(* IEC 61131-3 sources: kns-port-domestic/upstream/plc-process-lib/src/POUs/Control/FB_PID, 12 files *)

(* ---- FB_PID.decl.st ---- *)
// Назначение: ПИД-регулятор в идеальной форме (Kp, Ti, Td): D по измерению с фильтром первого
//             порядка, anti-windup обратным расчётом с постоянной слежения Tt (по своему выходу
//             или по фактическому выходу механизма rOutAct_pct), пределы и ограничение скорости
//             выхода, Manual и слежение (xTrack) с безударным переходом, внешнее или операторское
//             задание с рампой, прямое и обратное действие, зона нечувствительности, расчёт по
//             реальному dt источника времени и период расчёта tSample, реакция на недостоверную PV.
//             Внутреннее состояние (I, D, PV прошлого шага, задание после рампы, выход) — LREAL.
//             Режимы Auto, Manual, OutOfService (Local нет); одна тревога PvInvalid.
// Автор:      kr0nsch
// Версия:     0.1.0
// Документ:   docs/fb/FB_PID.md
FUNCTION_BLOCK FB_PID EXTENDS FB_DeviceBase
VAR_INPUT
    rPv_eu      : REAL;              // регулируемая величина, инж. ед.
    xPvValid    : BOOL;              // PV достоверна; по умолчанию FALSE — забытая привязка видна сразу
    xSpExt      : BOOL;              // задание от логики (каскад, график), а не от оператора
    rSpExt_eu   : REAL;              // внешнее задание, инж. ед.
    xTrack      : BOOL;              // слежение: выход := rTrack_pct (исполнительный механизм не в Auto)
    rTrack_pct  : REAL;              // значение для слежения, %
    rOutAct_pct : REAL;              // фактический выход механизма, % (при stCfg.xUseOutAct)
END_VAR
VAR_IN_OUT
    stCmd    : ST_PidCmd;            // команды HMI/SCADA; ФБ пишет слежение rSp_eu, rManualOut_pct
    stRetain : ST_DeviceRetain;      // используются eRemoteMode и xOutOfService
END_VAR
VAR_IN_OUT CONSTANT
    stCfg : ST_PidCfg;               // параметры (Persistent Variables приложения)
END_VAR
VAR_OUTPUT
    rOut_pct : REAL;                 // выход, %
    xSatHigh : BOOL;                 // выход на верхнем пределе rOutMax_pct
    xSatLow  : BOOL;                 // выход на нижнем пределе rOutMin_pct
    stSts    : ST_PidSts;            // состояние для HMI/SCADA
END_VAR
VAR
    stCfgLkg      : ST_PidCfg;       // последняя корректная конфигурация (LKG, нормативно)
    // --- состояние алгоритма (LREAL: малые приращения интегратора не теряются рядом с 50 %) ---
    lrOut_pct     : LREAL;           // выход u (он же u прошлого шага для ограничения скорости)
    lrI_pct       : LREAL;           // интегральная составляющая (после обновления этого шага)
    lrP_pct       : LREAL;           // пропорциональная составляющая последнего расчёта
    lrD_pct       : LREAL;           // дифференциальная составляющая последнего расчёта
    lrV_pct       : LREAL;           // v = P + I + D до ограничения, последний расчёт
    lrErr_pct     : LREAL;           // ошибка e' после зоны нечувствительности, % диапазона PV
    lrPvPrev_eu   : LREAL;           // PV прошлого расчёта (D по измерению)
    lrSp_eu       : LREAL;           // действующее задание (после рампы)
    lrSpTarget_eu : LREAL;           // цель задания после пределов (до рампы)
    lrDtCalc_s    : LREAL;           // dt последнего расчёта, с; 0 — шаг инициализации
    ltLastCalc    : LTIME;           // время последнего расчёта
    xCalcInit     : BOOL := TRUE;    // следующий расчёт — шаг инициализации (старт, PV вернулась, OOS)
    xFirstCalc    : BOOL := TRUE;    // расчёта ещё не было (первый расчёт ставит бит DT_GAP)
    xSpInit       : BOOL := TRUE;    // рампа задания не начата: первый расчёт берёт цель сразу
    // --- признаки последнего вызова (карта битов) ---
    xPvOk         : BOOL;            // xPvValid AND PV конечна
    xDtGap        : BOOL;            // разрыв времени: шаг инициализации этого вызова
    xSpInvalid    : BOOL;            // цель задания не конечна, удерживается прежняя
    xInDeadband   : BOOL;            // ошибка в зоне нечувствительности (последний расчёт)
    xOutRateLim   : BOOL;            // выход ограничен по скорости (последний расчёт в Auto)
    xTrackAct     : BOOL;            // выход следует за rTrack_pct
    xPvShed       : BOOL;            // ФБ сам перевёл контур в Manual по отказу PV (ShedToManual)
END_VAR
VAR_TEMP
    xAutoReq      : BOOL;            // в этом вызове запрошен Auto
    xHigherReq    : BOOL;            // запрошен Manual или OutOfService (старше Auto)
    eRes          : E_CmdResult;     // результат ProcessMode
    xSpTrack      : BOOL;            // задание следует за PV (Manual, xSpTrackPv)
    rSpRaw_eu     : REAL;            // цель задания до пределов
    xCalc         : BOOL;            // в этом вызове выполняется расчёт
    xInitStep     : BOOL;            // расчёт — шаг инициализации
    ltElapsed     : LTIME;           // время от последнего расчёта
    lrDt_s        : LREAL;           // шаг расчёта, с
    xPvFault      : BOOL;            // PV негодна в Auto без слежения: Failure
    eDevSt        : E_Ne107Status;   // вклад логики в NE 107
END_VAR

(* ---- CalcStep.method.decl.st ---- *)
// Шаг расчёта (контракт 17.4): рампа задания; ошибка со знаком действия в % диапазона PV; зона
// нечувствительности без скачка на границе (e' = e - DB·SIGN(e)); P = Kp·e'; D по измерению с
// фильтром Tf = Td/N (обратная разность Эйлера, устойчива при любом dt; в шаге инициализации
// D := 0); PV_prev := PV; v = P + I + D. Работает только с внутренним состоянием, stCfgLkg и
// входом rPv_eu (VAR_IN_OUT не трогает, R2)
METHOD PROTECTED CalcStep
VAR_INPUT
    xInit     : BOOL;    // шаг инициализации: D := 0
    lrStep_s  : LREAL;   // dt, с (0 в шаге инициализации)
    xSpFollow : BOOL;    // задание сразу равно цели (слежение задания за PV в Manual)
END_VAR
VAR
    lrPv_eu  : LREAL;    // PV этого вызова
    lrSign   : LREAL;    // +1 обратное действие, -1 прямое
    lrScale  : LREAL;    // % диапазона PV на инж. ед.
    lrE_pct  : LREAL;    // ошибка до зоны нечувствительности
    lrDb_pct : LREAL;    // зона нечувствительности
    lrKp     : LREAL;    // Kp
    lrTd_s   : LREAL;    // Td
    lrTf_s   : LREAL;    // постоянная фильтра Д: Td / N
END_VAR

(* ---- CalcStep.method.impl.st ---- *)
lrPv_eu := REAL_TO_LREAL(rPv_eu);
// рампа задания; первый расчёт и слежение за PV берут цель сразу
IF xSpInit OR xSpFollow THEN
    lrSp_eu := lrSpTarget_eu;
    xSpInit := FALSE;
ELSE
    lrSp_eu := RateStep(lrCurrent := lrSp_eu, lrTarget := lrSpTarget_eu,
                        lrRate := REAL_TO_LREAL(stCfgLkg.rSpRate_ups), lrStep_s := lrStep_s);
END_IF
// ошибка со знаком действия, % диапазона PV
IF stCfgLkg.eAction = E_PidAction.Direct THEN
    lrSign := -1.0;
ELSE
    lrSign := 1.0;
END_IF
lrScale := REAL_TO_LREAL(GVL_Const.PCT_FULL)
           / (REAL_TO_LREAL(stCfgLkg.rPvMax_eu) - REAL_TO_LREAL(stCfgLkg.rPvMin_eu));
lrE_pct := lrSign * (lrSp_eu - lrPv_eu) * lrScale;
// зона нечувствительности
lrDb_pct := REAL_TO_LREAL(stCfgLkg.rDeadband_pct);
xInDeadband := lrDb_pct > 0.0 AND ABS(lrE_pct) <= lrDb_pct;
IF ABS(lrE_pct) <= lrDb_pct THEN
    lrErr_pct := 0.0;
ELSIF lrE_pct > 0.0 THEN
    lrErr_pct := lrE_pct - lrDb_pct;
ELSE
    lrErr_pct := lrE_pct + lrDb_pct;
END_IF
// P по ошибке, D по измерению
lrKp := REAL_TO_LREAL(stCfgLkg.rKp);
lrP_pct := lrKp * lrErr_pct;
lrTd_s := REAL_TO_LREAL(stCfgLkg.rTd_s);
IF lrTd_s > 0.0 AND NOT xInit THEN
    lrTf_s := lrTd_s / REAL_TO_LREAL(stCfgLkg.rDFilterN);
    lrD_pct := lrTf_s / (lrTf_s + lrStep_s) * lrD_pct
               - lrKp * lrTd_s / (lrTf_s + lrStep_s) * lrSign * (lrPv_eu - lrPvPrev_eu) * lrScale;
ELSE
    lrD_pct := 0.0;
END_IF
lrPvPrev_eu := lrPv_eu;
lrV_pct := lrP_pct + lrI_pct + lrD_pct;

(* ---- CheckConfig.method.decl.st ---- *)
// Проверка конфигурации: биты wCfgErr (карта битов docs/fb/FB_PID.md). Неконечное значение
// REAL-параметра даёт бит его группы. Только считает, ничего не меняет
METHOD PROTECTED CheckConfig : WORD
VAR_IN_OUT CONSTANT
    stCfgIn : ST_PidCfg;   // проверяемая конфигурация
END_VAR
VAR
    wErr : WORD;           // непройденные проверки
END_VAR

(* ---- CheckConfig.method.impl.st ---- *)
// бит 0: действие — значение перечисления (сравнениями: строгое перечисление, L4 контракта)
IF stCfgIn.eAction <> E_PidAction.Reverse AND stCfgIn.eAction <> E_PidAction.Direct THEN
    wErr := wErr OR GVL_Const.PID_CFG_ACTION;
END_IF
// бит 1: Kp > 0
IF NOT F_IsFinite(rIn := stCfgIn.rKp) OR stCfgIn.rKp <= 0.0 THEN
    wErr := wErr OR GVL_Const.PID_CFG_KP;
END_IF
// бит 2: Ti >= 0, Td >= 0
IF NOT F_IsFinite(rIn := stCfgIn.rTi_s) OR NOT F_IsFinite(rIn := stCfgIn.rTd_s)
   OR stCfgIn.rTi_s < 0.0 OR stCfgIn.rTd_s < 0.0
THEN
    wErr := wErr OR GVL_Const.PID_CFG_TI_TD;
END_IF
// бит 3: фильтр Д — N в PID_DFILTER_N_MIN…MAX при Td > 0; неконечное N — всегда ошибка
IF NOT F_IsFinite(rIn := stCfgIn.rDFilterN)
   OR (stCfgIn.rTd_s > 0.0 AND (stCfgIn.rDFilterN < GVL_Const.PID_DFILTER_N_MIN
                                OR stCfgIn.rDFilterN > GVL_Const.PID_DFILTER_N_MAX))
THEN
    wErr := wErr OR GVL_Const.PID_CFG_DFILTER;
END_IF
// бит 4: Tt >= 0 (0 — авто)
IF NOT F_IsFinite(rIn := stCfgIn.rTt_s) OR stCfgIn.rTt_s < 0.0 THEN
    wErr := wErr OR GVL_Const.PID_CFG_TT;
END_IF
// бит 5: диапазон PV
IF NOT F_IsFinite(rIn := stCfgIn.rPvMin_eu) OR NOT F_IsFinite(rIn := stCfgIn.rPvMax_eu)
   OR stCfgIn.rPvMin_eu >= stCfgIn.rPvMax_eu
THEN
    wErr := wErr OR GVL_Const.PID_CFG_PV_RANGE;
END_IF
// бит 6: пределы задания (равные допустимы — задание фиксировано)
IF NOT F_IsFinite(rIn := stCfgIn.rSpMin_eu) OR NOT F_IsFinite(rIn := stCfgIn.rSpMax_eu)
   OR stCfgIn.rSpMin_eu > stCfgIn.rSpMax_eu
THEN
    wErr := wErr OR GVL_Const.PID_CFG_SP_RANGE;
END_IF
// бит 7: пределы выхода в 0…100 %, min < max
IF NOT F_IsFinite(rIn := stCfgIn.rOutMin_pct) OR NOT F_IsFinite(rIn := stCfgIn.rOutMax_pct)
   OR stCfgIn.rOutMin_pct < 0.0 OR stCfgIn.rOutMax_pct > GVL_Const.PCT_FULL
   OR stCfgIn.rOutMin_pct >= stCfgIn.rOutMax_pct
THEN
    wErr := wErr OR GVL_Const.PID_CFG_OUT_RANGE;
END_IF
// бит 8: зона нечувствительности в 0…PID_DEADBAND_MAX_PCT
IF NOT F_IsFinite(rIn := stCfgIn.rDeadband_pct) OR stCfgIn.rDeadband_pct < 0.0
   OR stCfgIn.rDeadband_pct > GVL_Const.PID_DEADBAND_MAX_PCT
THEN
    wErr := wErr OR GVL_Const.PID_CFG_DEADBAND;
END_IF
// бит 9: скорости рампы задания и выхода >= 0 (0 — без ограничения)
IF NOT F_IsFinite(rIn := stCfgIn.rSpRate_ups) OR NOT F_IsFinite(rIn := stCfgIn.rOutRate_pctps)
   OR stCfgIn.rSpRate_ups < 0.0 OR stCfgIn.rOutRate_pctps < 0.0
THEN
    wErr := wErr OR GVL_Const.PID_CFG_RATES;
END_IF
// бит 10: tDtMax > 0, tSample < tDtMax
IF stCfgIn.tDtMax = T#0S OR stCfgIn.tSample >= stCfgIn.tDtMax THEN
    wErr := wErr OR GVL_Const.PID_CFG_SAMPLE;
END_IF
// бит 11: реакция на отказ PV — значение перечисления; безопасный выход в пределах выхода
IF (stCfgIn.ePvFailAction <> E_PidPvFailAction.Hold AND stCfgIn.ePvFailAction <> E_PidPvFailAction.SafeOut
    AND stCfgIn.ePvFailAction <> E_PidPvFailAction.ShedToManual)
   OR NOT F_IsFinite(rIn := stCfgIn.rSafeOut_pct)
   OR stCfgIn.rSafeOut_pct < stCfgIn.rOutMin_pct OR stCfgIn.rSafeOut_pct > stCfgIn.rOutMax_pct
THEN
    wErr := wErr OR GVL_Const.PID_CFG_PV_FAIL;
END_IF
// бит 12: приоритеты тревог — значения перечисления
IF NOT CheckAlarmCfg(astCfg := stCfgIn.astAlarm) THEN
    wErr := wErr OR GVL_Const.PID_CFG_ALARM;
END_IF
CheckConfig := wErr;

(* ---- FB_PID.impl.st ---- *)
// 0. Первый вызов: число слотов тревог и тип устройства (до ProcessMode)
IF xFirstCall THEN
    uiAlarmCount := GVL_Const.PID_ALARM_COUNT;
    eDevType := E_DeviceType.Pid;
END_IF

// 1. Время
BeginCycle();

// 2. Конфигурация (LKG); достоверность PV
IF AcceptCfg(wErr := CheckConfig(stCfgIn := stCfg)) THEN
    stCfgLkg := stCfg;
END_IF
xPvOk := xPvValid AND F_IsFinite(rIn := rPv_eu);
// 2а. Старт ПЛК: выход — фактический выход механизма: rOutAct_pct при xUseOutAct, иначе
//     rTrack_pct при слежении, иначе stCmd.rManualOut_pct. Интегратор инициализирует шаг
//     инициализации первого расчёта (I := u - P)
IF xFirstCall THEN
    IF stCfgLkg.xUseOutAct AND F_IsFinite(rIn := rOutAct_pct) THEN
        lrOut_pct := REAL_TO_LREAL(rOutAct_pct);
    ELSIF xTrack AND F_IsFinite(rIn := rTrack_pct) THEN
        lrOut_pct := REAL_TO_LREAL(rTrack_pct);
    ELSIF F_IsFinite(rIn := stCmd.rManualOut_pct) THEN
        lrOut_pct := REAL_TO_LREAL(stCmd.rManualOut_pct);
    END_IF
END_IF

// 3. Reset: фиксируемых отказов у ПИД нет — команда принимается (тревоги квитирует RunAlarms)
IF xResetReq OR stCmd.stCommon.xReset THEN
    SetCmdResult(eResult := E_CmdResult.Accepted);
END_IF

// 4. Режим. Запрос Auto без корректной Cfg (RejectedCfg) или при негодной PV (RejectedFault)
//    снимается до ProcessMode. Если в том же вызове есть старший запрос (Manual, OutOfService),
//    Auto снимается молча: ProcessMode обработает старший как одну команду
xAutoReq := stCmd.stCommon.xSetAuto OR (xModeReq AND eModeReq = E_DeviceMode.Auto);
xHigherReq := stCmd.stCommon.xSetOos OR stCmd.stCommon.xSetManual
              OR (xModeReq AND eModeReq <> E_DeviceMode.Auto);
IF xAutoReq AND (NOT xCfgEverOk OR NOT xPvOk) THEN
    IF NOT xHigherReq THEN
        IF NOT xCfgEverOk THEN
            SetCmdResult(eResult := E_CmdResult.RejectedCfg);
        ELSE
            SetCmdResult(eResult := E_CmdResult.RejectedFault);
        END_IF
    END_IF
    stCmd.stCommon.xSetAuto := FALSE;
    IF eModeReq = E_DeviceMode.Auto THEN
        xModeReq := FALSE;
    END_IF
END_IF
eRes := ProcessMode(xLocalSel := FALSE, xLocalSupported := FALSE, xOosAllowed := TRUE,
                    stCmd := stCmd.stCommon, stRetain := stRetain);
IF eRes <> E_CmdResult.None THEN
    SetCmdResult(eResult := eRes);
END_IF

// 5. Переходы логики: PV негодна в Auto без слежения и реакция ShedToManual — в Manual с
//    текущим выходом (stCmd.rManualOut_pct уже равен выходу: слежение в Auto). Признак
//    сброса держит тревогу PvInvalid в Manual, пока PV негодна; снимают его годная PV и
//    выбор оператором OutOfService (docs/fb/FB_PID.md, P-15)
IF xCfgEverOk AND eMode = E_DeviceMode.Auto AND NOT xPvOk AND NOT xTrack
   AND stCfgLkg.ePvFailAction = E_PidPvFailAction.ShedToManual
THEN
    SwitchRemoteMode(eNew := E_DeviceMode.Manual, stRetain := stRetain);
    xPvShed := TRUE;
END_IF
IF xPvOk OR eMode <> E_DeviceMode.Manual THEN
    xPvShed := FALSE;
END_IF

// 6. Логика по stCfgLkg
// 6.1 Задание: цель (внешнее, PV при слежении задания в Manual или операторское), пределы.
//     Неконечная цель — прежняя цель и предупреждение; пределы действуют и на неё (NaN с
//     первого вызова, смена пределов при NaN; P-16). Внешнее задание и PV пишутся в
//     stCmd.rSp_eu: переход на операторское задание без рывка
xSpTrack := eMode = E_DeviceMode.Manual AND stCfgLkg.xSpTrackPv AND NOT xSpExt AND xPvOk;
IF xSpExt THEN
    rSpRaw_eu := rSpExt_eu;
ELSIF xSpTrack THEN
    rSpRaw_eu := rPv_eu;
ELSE
    rSpRaw_eu := stCmd.rSp_eu;
END_IF
xSpInvalid := NOT F_IsFinite(rIn := rSpRaw_eu);
IF NOT xSpInvalid THEN
    lrSpTarget_eu := REAL_TO_LREAL(rSpRaw_eu);
    IF xCfgEverOk AND (xSpExt OR xSpTrack) THEN
        stCmd.rSp_eu := rSpRaw_eu;
    END_IF
END_IF
lrSpTarget_eu := LIMIT(REAL_TO_LREAL(stCfgLkg.rSpMin_eu), lrSpTarget_eu, REAL_TO_LREAL(stCfgLkg.rSpMax_eu));

// 6.2 Нужен ли расчёт. Без корректной Cfg и при негодной PV расчёта нет, следующий — шаг
//     инициализации; в OutOfService расчёта нет (выход из OOS ставит инициализацию в хуке).
//     LTIME без знака: «время назад» проверяется до вычитания. Разрыв больше tDtMax и «время
//     назад» — шаг инициализации с битом DT_GAP; dt = 0 — расчёта нет
xCalc := FALSE;
xInitStep := FALSE;
xDtGap := FALSE;
lrDt_s := 0.0;
IF NOT xCfgEverOk OR NOT xPvOk THEN
    xCalcInit := TRUE;
ELSIF eMode <> E_DeviceMode.OutOfService THEN
    IF xCalcInit OR ltNow < ltLastCalc THEN
        xCalc := TRUE;
        xInitStep := TRUE;
        xDtGap := xFirstCalc OR NOT xCalcInit;
    ELSE
        ltElapsed := ltNow - ltLastCalc;
        IF ltElapsed > TIME_TO_LTIME(stCfgLkg.tDtMax) THEN
            xCalc := TRUE;
            xInitStep := TRUE;
            xDtGap := TRUE;
        ELSIF ltElapsed > LTIME#0S AND ltElapsed >= TIME_TO_LTIME(stCfgLkg.tSample) THEN
            xCalc := TRUE;
            lrDt_s := F_LTimeToSec(ltIn := ltElapsed);
        END_IF
    END_IF
END_IF

// 6.3 Шаг расчёта (контракт 17.4): рампа задания, ошибка, зона нечувствительности, P, D, v
IF xCalc THEN
    ltLastCalc := ltNow;
    xCalcInit := FALSE;
    xFirstCalc := FALSE;
    lrDtCalc_s := lrDt_s;
    CalcStep(xInit := xInitStep, lrStep_s := lrDt_s, xSpFollow := xSpTrack);
END_IF

// 6.4 Выход по старшинству (контракт 2.6, 17.5), интегратор, rOut_pct, xSatHigh, xSatLow
SelectOutput(xCalcNow := xCalc, xInit := xInitStep, lrStep_s := lrDt_s, rManualOut_pct := stCmd.rManualOut_pct);

// 6.5 Слежение в Cmd: в Auto, OutOfService и при слежении выход пишется в rManualOut_pct
IF xCfgEverOk AND (eMode <> E_DeviceMode.Manual OR xTrackAct) THEN
    stCmd.rManualOut_pct := LREAL_TO_REAL(lrOut_pct);
END_IF

// 7. Тревоги: слот 0 PvInvalid — PV негодна в Auto или после сброса в Manual по отказу PV
axAlmCond[E_PidAlarm.PvInvalid] := NOT xPvOk AND (eMode = E_DeviceMode.Auto OR xPvShed);
axAlmSuppress[E_PidAlarm.PvInvalid] := FALSE;
arAlmValue[E_PidAlarm.PvInvalid] := SEL(F_IsFinite(rIn := rPv_eu), 0.0, rPv_eu);
RunAlarms(udiIdBase := stCfgLkg.udiAlarmIdBase, stCmd := stCmd.stCommon, astCfg := stCfgLkg.astAlarm);

// 8. Состояние
xPvFault := NOT xPvOk AND eMode = E_DeviceMode.Auto AND NOT xTrack;
IF xPvFault THEN
    eDevSt := E_Ne107Status.Failure;
ELSE
    eDevSt := E_Ne107Status.Good;
END_IF
stSts.rSpTarget_eu := LREAL_TO_REAL(lrSpTarget_eu);
stSts.rSp_eu := LREAL_TO_REAL(lrSp_eu);
stSts.rPv_eu := SEL(F_IsFinite(rIn := rPv_eu), 0.0, rPv_eu);   // NaN из Modbus — 0.0 (R6), PV_FAIL в битах
stSts.rErr_pct := LREAL_TO_REAL(lrErr_pct);
stSts.rOut_pct := rOut_pct;
stSts.rP_pct := LREAL_TO_REAL(lrP_pct);
stSts.rI_pct := LREAL_TO_REAL(lrI_pct);
stSts.rD_pct := LREAL_TO_REAL(lrD_pct);
stSts.rDt_ms := LREAL_TO_REAL(lrDtCalc_s * GVL_Const.MS_PER_S);
FinishCycle(eDevStatus := eDevSt,
            xAvailableDev := eMode = E_DeviceMode.Auto AND xPvOk AND NOT xTrack,
            wLow := SEL(xSatHigh, 0, GVL_Const.PID_STS_SAT_HIGH)
                    OR SEL(xSatLow, 0, GVL_Const.PID_STS_SAT_LOW)
                    OR SEL(xCfgEverOk AND NOT xSpInit AND eMode <> E_DeviceMode.OutOfService
                           AND lrSp_eu <> lrSpTarget_eu, 0, GVL_Const.PID_STS_SP_RAMPING)
                    OR SEL(xInDeadband, 0, GVL_Const.PID_STS_IN_DEADBAND)
                    OR SEL(xPvOk, GVL_Const.PID_STS_PV_FAIL, 0)            // бит при PV негодна
                    OR SEL(xDtGap, 0, GVL_Const.PID_STS_DT_GAP)
                    OR SEL(xTrackAct, 0, GVL_Const.PID_STS_TRACKING)
                    OR SEL(xOutRateLim, 0, GVL_Const.PID_STS_OUT_RATE_LIMITED),
            wFaultBits := SEL(xPvFault, 0, GVL_Const.PID_FLT_PV_INVALID),
            wWarnBits := SEL(xDtGap, 0, GVL_Const.PID_WRN_DT_GAP) OR SEL(xSpInvalid, 0, GVL_Const.PID_WRN_SP_INVALID),
            stCommon := stSts.stCommon);

(* ---- OnModeChanged.method.decl.st ---- *)
// Хук смены режима: сначала база (SUPER^). Выход из OutOfService — следующий расчёт будет шагом
// инициализации (PV_prev := PV, D := 0, I := u - P): за время OOS PV и время ушли. Вход в Auto —
// предустановка I := u - P - D по последнему расчёту: v = u, переход без рывка (в Manual и при
// слежении тело держит это равенство каждый вызов). VAR_IN_OUT устройства не трогает (R2)
METHOD PROTECTED OnModeChanged
VAR_INPUT
    eOld : E_DeviceMode;   // режим до смены
    eNew : E_DeviceMode;   // новый режим
END_VAR

(* ---- OnModeChanged.method.impl.st ---- *)
SUPER^.OnModeChanged(eOld := eOld, eNew := eNew);
IF eOld = E_DeviceMode.OutOfService THEN
    xCalcInit := TRUE;
END_IF
IF eNew = E_DeviceMode.Auto THEN
    lrI_pct := lrOut_pct - lrP_pct - lrD_pct;
END_IF

(* ---- RateStep.method.decl.st ---- *)
// Ограничение скорости в LREAL (рампа задания и ограничение скорости выхода): значение движется
// от lrCurrent к lrTarget не быстрее lrRate ед./с за шаг lrStep_s. Скорость <= 0 — сразу к
// цели (в том числе в шаге инициализации); шаг <= 0 при заданной скорости — без изменения.
// F_RateLimit не подходит: вход и результат REAL, приращения рампы меньше шага REAL теряются
METHOD PROTECTED RateStep : LREAL
VAR_INPUT
    lrCurrent : LREAL;   // текущее значение
    lrTarget  : LREAL;   // цель
    lrRate    : LREAL;   // предел скорости, ед./с; <= 0 — без ограничения
    lrStep_s  : LREAL;   // шаг времени, с
END_VAR

(* ---- RateStep.method.impl.st ---- *)
IF lrRate <= 0.0 THEN
    RateStep := lrTarget;
ELSIF lrStep_s <= 0.0 THEN
    RateStep := lrCurrent;
ELSIF lrTarget > lrCurrent THEN
    RateStep := MIN(lrTarget, lrCurrent + lrRate * lrStep_s);
ELSE
    RateStep := MAX(lrTarget, lrCurrent - lrRate * lrStep_s);
END_IF

(* ---- SelectOutput.method.decl.st ---- *)
// Выход по старшинству (контракт 2.6, 17.5): нет корректной Cfg > OutOfService > слежение >
// Manual > Auto с негодной PV > Auto. Вне Auto интегратор предустанавливается I := u - P - D (при
// возврате в Auto v = u, рывка нет). Auto: пределы, ограничение скорости, обратный расчёт
// I += Kp·dt/Ti·e' + MIN(dt/Tt, 1)·(u_aw - v), u_aw — выход ФБ или rOutAct_pct (xUseOutAct).
// Пишет rOut_pct, xSatHigh, xSatLow. Значение оператора — параметром (VAR_IN_OUT не трогает, R2)
METHOD PROTECTED SelectOutput
VAR_INPUT
    xCalcNow       : BOOL;    // в этом вызове был расчёт (CalcStep)
    xInit          : BOOL;    // расчёт — шаг инициализации
    lrStep_s       : LREAL;   // dt расчёта, с
    rManualOut_pct : REAL;    // stCmd.rManualOut_pct: выход оператора
END_VAR
VAR
    lrOutMin_pct : LREAL;     // нижний предел выхода
    lrOutMax_pct : LREAL;     // верхний предел выхода
    lrULim_pct   : LREAL;     // LIMIT(OutMin, v, OutMax)
    lrUAw_pct    : LREAL;     // выход для обратного расчёта (u или rOutAct_pct)
    lrKp         : LREAL;     // Kp
    lrTi_s       : LREAL;     // Ti
    lrTd_s       : LREAL;     // Td
    lrTt_s       : LREAL;     // постоянная слежения anti-windup
END_VAR

(* ---- SelectOutput.method.impl.st ---- *)
lrOutMin_pct := REAL_TO_LREAL(stCfgLkg.rOutMin_pct);
lrOutMax_pct := REAL_TO_LREAL(stCfgLkg.rOutMax_pct);
xTrackAct := FALSE;
IF NOT xCfgEverOk THEN
    // расчёта нет: выход от оператора в пределах 0…100 %; неконечное значение — выход прежний
    IF F_IsFinite(rIn := rManualOut_pct) THEN
        lrOut_pct := LIMIT(0.0, REAL_TO_LREAL(rManualOut_pct), REAL_TO_LREAL(GVL_Const.PCT_FULL));
    END_IF
    xOutRateLim := FALSE;
ELSIF eMode = E_DeviceMode.OutOfService THEN
    // выход удерживается, расчёта нет
    lrI_pct := lrOut_pct - lrP_pct - lrD_pct;
    xOutRateLim := FALSE;
ELSIF xTrack THEN
    // слежение: без пределов (механизм может стоять на 0); неконечное значение — выход прежний
    xTrackAct := TRUE;
    IF F_IsFinite(rIn := rTrack_pct) THEN
        lrOut_pct := REAL_TO_LREAL(rTrack_pct);
    END_IF
    lrI_pct := lrOut_pct - lrP_pct - lrD_pct;
    xOutRateLim := FALSE;
ELSIF eMode = E_DeviceMode.Manual THEN
    IF F_IsFinite(rIn := rManualOut_pct) THEN
        lrOut_pct := LIMIT(lrOutMin_pct, REAL_TO_LREAL(rManualOut_pct), lrOutMax_pct);
    END_IF
    lrI_pct := lrOut_pct - lrP_pct - lrD_pct;
    xOutRateLim := FALSE;
ELSIF NOT xPvOk THEN
    // Auto, PV негодна: Hold — выход удерживается, SafeOut — rSafeOut_pct; интегратор заморожен,
    // возврат PV — шаг инициализации (I := u - P): без рывка
    IF stCfgLkg.ePvFailAction = E_PidPvFailAction.SafeOut THEN
        lrOut_pct := REAL_TO_LREAL(stCfgLkg.rSafeOut_pct);
    END_IF
    xOutRateLim := FALSE;
ELSIF xCalcNow AND xInit THEN
    // шаг инициализации: выход прежний, интегрирования нет
    lrI_pct := lrOut_pct - lrP_pct - lrD_pct;
    xOutRateLim := FALSE;
ELSIF xCalcNow THEN
    // Auto: пределы, ограничение скорости, обратный расчёт по u или по rOutAct_pct
    lrULim_pct := LIMIT(lrOutMin_pct, lrV_pct, lrOutMax_pct);
    lrOut_pct := RateStep(lrCurrent := lrOut_pct, lrTarget := lrULim_pct,
                          lrRate := REAL_TO_LREAL(stCfgLkg.rOutRate_pctps), lrStep_s := lrStep_s);
    xOutRateLim := lrOut_pct <> lrULim_pct;
    IF stCfgLkg.xUseOutAct AND F_IsFinite(rIn := rOutAct_pct) THEN
        lrUAw_pct := REAL_TO_LREAL(rOutAct_pct);
    ELSE
        lrUAw_pct := lrOut_pct;
    END_IF
    lrKp := REAL_TO_LREAL(stCfgLkg.rKp);
    lrTi_s := REAL_TO_LREAL(stCfgLkg.rTi_s);
    lrTd_s := REAL_TO_LREAL(stCfgLkg.rTd_s);
    IF lrTi_s > 0.0 THEN
        // Tt: rTt_s, если задана; иначе SQRT(Ti·Td) при Td > 0; иначе Ti
        IF stCfgLkg.rTt_s > 0.0 THEN
            lrTt_s := REAL_TO_LREAL(stCfgLkg.rTt_s);
        ELSIF lrTd_s > 0.0 THEN
            lrTt_s := SQRT(lrTi_s * lrTd_s);
        ELSE
            lrTt_s := lrTi_s;
        END_IF
        lrI_pct := lrI_pct + lrKp * lrStep_s / lrTi_s * lrErr_pct
                   + MIN(lrStep_s / lrTt_s, 1.0) * (lrUAw_pct - lrV_pct);
    END_IF
END_IF
rOut_pct := LREAL_TO_REAL(lrOut_pct);
xSatHigh := xCfgEverOk AND lrOut_pct >= lrOutMax_pct;
xSatLow := xCfgEverOk AND lrOut_pct <= lrOutMin_pct;
